// TIA Portal V20 export
// export: Created 2026-10-11T05:25:30.5137323Z, ExportSetting WithDefaults, DisplayName Totally Integrated Automation Portal, DisplayVersion V20, DisplayName TIA Portal Openness, DisplayVersion V20, DisplayName TIA Portal Teamcenter Gateway, DisplayVersion V20, DisplayName TIA Portal Version Control Interface, DisplayVersion V20, DisplayName SINAMICS Startdrive Advanced, DisplayVersion V20 SP1 Update 2, DisplayName SINAMICS Startdrive G110M, G120, G120C, G120D, G120P, G115D, DisplayVersion V20 SP1 Update 2, DisplayName SINAMICS Startdrive G130, G150, S120, S150, SINAMICS MV, G220, S200, S210, DisplayVersion V20 SP1 Update 2, DisplayName STEP 7 Professional, DisplayVersion V20, DisplayName STEP 7 Safety, DisplayVersion V20, DisplayName WinCC Basic/Comfort/Advanced, DisplayVersion V20, DisplayName WinCC Professional, DisplayVersion V20, DisplayName WinCC Unified, DisplayVersion V20
FUNCTION "FRK_AccessFinish" : Void   // FC34, SCL
{ S7_Optimized_Access := 'TRUE' }
VERSION : 0.1
// stored: AutoNumber true, IsIECCheckEnabled false, SetENOAutomatically false, UDAEnableTagReadback false
   VAR_INPUT
      Unit : "FRK_Unit";
      Response : "ST_HmiResponse";
      SourcePath : WString;
   END_VAR
   VAR_IN_OUT
      Access : "FRK_Access";
      History : Array[1..16] of "ST_Diagnostic";
      Head : Int;
      Revision : UDInt;
   END_VAR
   VAR_TEMP
      What : WString[160];
      AuditPath : WString[255];
   END_VAR
BEGIN

   IF NOT #Unit.RequestPending THEN
       RETURN;
   END_IF;
   CASE #Unit.Request.Kind OF
       23, 15,
       16, 17,
       1:
           RETURN;
       2:
           "FRK_AccessAudit"(History := #History,
                             Head := #Head,
                             What := WSTRING#'std.audit.logout',
                             Who := #Unit.RequestUser,
                             SourcePath := #SourcePath);
           #Revision := "FRK_ConfigRevision"(Previous := #Revision);
           RETURN;
       ELSE
           #What := WSTRING#'std.audit.accessDenied';
   END_CASE;
   IF #Response.Accepted THEN
       #What := WSTRING#'std.audit.operatorMutation';
       IF #Access.CurrentLevel > 0 THEN
           #Access.LastActivity := "FRK_Clock".NowMs;
       END_IF;
       IF #Unit.Request.Kind = 24 THEN
           #Revision := "FRK_ConfigRevision"(Previous := #Revision);
       END_IF;
   END_IF;
   #AuditPath := #SourcePath;
   IF #Unit.Request.Kind = 11 THEN
       #AuditPath := #Unit.Request.TargetPath;
       IF #Response.Accepted THEN
           #What := WSTRING#'std.audit.manualCommandAccepted';
       ELSE
           #What := WSTRING#'std.audit.manualCommandRejected';
       END_IF;
   END_IF;
   #What := CONCAT(IN1 := #What, IN2 := WSTRING#' kind=');
   #What := CONCAT(IN1 := #What, IN2 := DINT_TO_WSTRING(#Unit.Request.Kind));
   #What := CONCAT(IN1 := #What, IN2 := WSTRING#' value=');
   #What := CONCAT(IN1 := #What, IN2 := DINT_TO_WSTRING(#Unit.Request.IntValue));
   "FRK_AccessAudit"(History := #History,
                     Head := #Head,
                     What := #What,
                     Who := #Unit.RequestUser,
                     SourcePath := #AuditPath);
END_FUNCTION
